// TIA Portal V20 export
Screen "Pop-up_EEM_LEGEND_Popup"  430x496
  ScreenItem "Background" at 0,0 size 430x496  Type=HmiRectangle
  ScreenItem "Text_Legend1" at 1,1 size 428x25  Type=HmiTextBox
  ScreenItem "Text_Legend2" at 10,32 size 325x20  Type=HmiTextBox
  ScreenItem "Text_ButtonsLeds" at 10,56 size 150x20  Type=HmiTextBox
  ScreenItem "Cancel Mode" at 337,3 size 90x60  Type=HmiButton
  ScreenItem "Text_P-Meas1" at 10,78 size 60x40  Type=HmiTextBox
  ScreenItem "Text_P-Meas2" at 75,76 size 350x54  Type=HmiTextBox
  ScreenItem "Text_Control+1" at 10,190 size 60x40  Type=HmiTextBox
  ScreenItem "Text_UIPE1" at 10,232 size 60x40  Type=HmiTextBox
  ScreenItem "Symbol_Meas1" at 0,0 size 100x30  Type=HmiCircle
  ScreenItem "Symbol_RefMeas1" at 0,0 size 100x30  Type=HmiCircle
  ScreenItem "Symbol1_RefMeas1" at 0,0 size 100x30  Type=HmiCircle
  ScreenItem "Text_Meas2" at 75,132 size 350x18  Type=HmiTextBox
  ScreenItem "Text_RefMeas2" at 75,151 size 350x18  Type=HmiTextBox
  ScreenItem "Text_DevNo_3" at 75,170 size 350x18  Type=HmiTextBox
  ScreenItem "Text_Control+2" at 75,193 size 350x35  Type=HmiTextBox
  ScreenItem "Button_ResetText_4" at 75,235 size 350x35  Type=HmiTextBox
  ScreenItem "Text_InfoMachine1" at 10,274 size 60x40  Type=HmiTextBox
  ScreenItem "Symbol2_RefMeas1" at 0,0 size 100x30  Type=HmiCircle
  ScreenItem "Text_InfoMachine2" at 75,277 size 350x35  Type=HmiTextBox
  ScreenItem "Text_ScreenContent" at 10,318 size 150x20  Type=HmiTextBox
  ScreenItem "Text_MeasPoint" at 10,340 size 415x35  Type=HmiTextBox
  ScreenItem "Symbol3_RefMeas1" at 0,0 size 100x30  Type=HmiCircle
  ScreenItem "Text_GraphDisplay1" at 10,377 size 415x35  Type=HmiTextBox
  ScreenItem "Text_GraphDisplay2" at 10,414 size 415x35  Type=HmiTextBox
  ScreenItem "Text_GraphDisplay3" at 10,451 size 415x35  Type=HmiTextBox
